(* IEC 61131-3 sources: plc-iiot-stack/tests/POUs/FB_MqttAlarms_Test, 12 files *)

(* ---- BudgetAndDisabledPriority.method.decl.st ---- *)
// Не больше uiMaxPerCycle за вызов; приоритет None — тревога пропускается.
METHOD PRIVATE BudgetAndDisabledPriority
VAR_INST
    fbFake : FB_MqttClientFake;
    fbAlm : FB_MqttAlarms;
    aAlm : ARRAY[1..3] OF ST_IiotAlarm;
    aWords : ARRAY[1..2] OF ST_IiotAlarmWords;
END_VAR

(* ---- ChangeWhileOfflineIsEventAfterReconnect.method.decl.st ---- *)
// Тревога сработала, пока связи не было: после переподключения — событие с текущим ts и prev_state
// последней публикации.
METHOD PRIVATE ChangeWhileOfflineIsEventAfterReconnect
VAR_INST
    fbFake : FB_MqttClientFake;
    fbAlm : FB_MqttAlarms;
    aAlm : ARRAY[1..3] OF ST_IiotAlarm;
    aWords : ARRAY[1..2] OF ST_IiotAlarmWords;
END_VAR

(* ---- EventsFollowWordChanges.method.decl.st ---- *)
// Появление, квитирование, снятие: Activated, Acked, Cleared.
METHOD PRIVATE EventsFollowWordChanges
VAR_INST
    fbFake : FB_MqttClientFake;
    fbAlm : FB_MqttAlarms;
    aAlm : ARRAY[1..3] OF ST_IiotAlarm;
    aWords : ARRAY[1..2] OF ST_IiotAlarmWords;
END_VAR

(* ---- ReconnectRepeatsLastEventWithItsTs.method.decl.st ---- *)
// Тревога сработала, связь пропала и вернулась: событие Activated повторяется с исходными ts и prev_state
// (в InfluxDB та же точка) — дашборды и отчёт не считают его вторым срабатыванием.
METHOD PRIVATE ReconnectRepeatsLastEventWithItsTs
VAR_INST
    fbFake : FB_MqttClientFake;
    fbAlm : FB_MqttAlarms;
    aAlm : ARRAY[1..3] OF ST_IiotAlarm;
    aWords : ARRAY[1..2] OF ST_IiotAlarmWords;
END_VAR

(* ---- ReturnUnackedThenAck.method.decl.st ---- *)
// Условие ушло без квитирования — RtnUnack/Cleared, затем квитирование — Normal/Acked.
METHOD PRIVATE ReturnUnackedThenAck
VAR_INST
    fbFake : FB_MqttClientFake;
    fbAlm : FB_MqttAlarms;
    aAlm : ARRAY[1..3] OF ST_IiotAlarm;
    aWords : ARRAY[1..2] OF ST_IiotAlarmWords;
END_VAR

(* ---- Setup.method.decl.st ---- *)
// Три тревоги: P101.FTS (слот 0, Medium) и P101.FTP (слот 2, High) — слова 1; LT101.HH (слот 0, High) — слова 2.
METHOD PRIVATE Setup
VAR_IN_OUT
    fbClient : FB_MqttClientFake;
    aAlarmTable : ARRAY[1..3] OF ST_IiotAlarm;
END_VAR

(* ---- ShelvedAndOutOfService.method.decl.st ---- *)
// Отложена/возвращена и вывод устройства из работы: Shelved, Unshelved, OosOn.
METHOD PRIVATE ShelvedAndOutOfService
VAR_INST
    fbFake : FB_MqttClientFake;
    fbAlm : FB_MqttAlarms;
    aAlm : ARRAY[1..3] OF ST_IiotAlarm;
    aWords : ARRAY[1..2] OF ST_IiotAlarmWords;
END_VAR

(* ---- SnapshotAfterBirthExactJson.method.decl.st ---- *)
// После рождения узла — снимок всех тревог; точный JSON, QoS 1, retain.
METHOD PRIVATE SnapshotAfterBirthExactJson
VAR_INST
    fbFake : FB_MqttClientFake;
    fbAlm : FB_MqttAlarms;
    aAlm : ARRAY[1..3] OF ST_IiotAlarm;
    aWords : ARRAY[1..2] OF ST_IiotAlarmWords;
END_VAR

(* ---- SnapshotAfterReconnectShowsCurrentState.method.decl.st ---- *)
// После переподключения — текущее состояние повтором первой публикации (снимка) с её ts, а не событие.
METHOD PRIVATE SnapshotAfterReconnectShowsCurrentState
VAR_INST
    fbFake : FB_MqttClientFake;
    fbAlm : FB_MqttAlarms;
    aAlm : ARRAY[1..3] OF ST_IiotAlarm;
    aWords : ARRAY[1..2] OF ST_IiotAlarmWords;
END_VAR

(* ---- StationAlarmIdAndLongSuffix.method.decl.st ---- *)
// Тревога станции флагмана KNS1.NOAUTO: номер 100009 (больше UINT), суффикс из шести знаков, бит slot - 1.
METHOD PRIVATE StationAlarmIdAndLongSuffix
VAR_INST
    fbFake : FB_MqttClientFake;
    fbAlm : FB_MqttAlarms;
    aAlm : ARRAY[1..1] OF ST_IiotAlarm;
    aWords : ARRAY[1..1] OF ST_IiotAlarmWords;
END_VAR

(* ---- SuppressedByDesignFromWords.method.decl.st ---- *)
// Бит wAlmSuppressed устройства (plc-process-lib 1.0) — состояние SuppressedByDesign и причины Suppressed/Unsuppressed.
METHOD PRIVATE SuppressedByDesignFromWords
VAR_INST
    fbFake : FB_MqttClientFake;
    fbAlm : FB_MqttAlarms;
    aAlm : ARRAY[1..3] OF ST_IiotAlarm;
    aWords : ARRAY[1..2] OF ST_IiotAlarmWords;
END_VAR

(* ---- WordsOutOfTableMeanNormal.method.decl.st ---- *)
// Строка слов вне таблицы — тревога в норме, без выхода за массив.
METHOD PRIVATE WordsOutOfTableMeanNormal
VAR_INST
    fbFake : FB_MqttClientFake;
    fbAlm : FB_MqttAlarms;
    aAlm : ARRAY[1..3] OF ST_IiotAlarm;
    aWords : ARRAY[1..2] OF ST_IiotAlarmWords;
END_VAR
